(* IEC 61131-3 sources: Lasal-MCP/examples/SampleSource/LASALScreenAdvancedSolution/LASALScreenAdvancedSolution/LASALScreenAdvacnedSolution/Stations/Terminal/HMI/Network/ValueNet, 1 file *)

(* ---- ONE_ValueNet_Table.st ---- *)
#define OBJECTS_CONFIG

FUNCTION GLOBAL TAB ONE_ValueNet
-1$UINT, 0$UINT,
0$UINT, 0$UINT,

1$UDINT,
TO_UDINT(443191026), "MyValues", 0$UINT, 0$UINT, 20$UINT,

_NO_ATTR, TO_UDINT(3497334281), "MYVALUES1",
_NO_ATTR, TO_UDINT(2379682451), "MYVALUES10",
_NO_ATTR, TO_UDINT(4207944197), "MYVALUES11",
_NO_ATTR, TO_UDINT(1675195327), "MYVALUES12",
_NO_ATTR, TO_UDINT(350110505), "MYVALUES13",
_NO_ATTR, TO_UDINT(2327500426), "MYVALUES14",
_NO_ATTR, TO_UDINT(4257080860), "MYVALUES15",
_NO_ATTR, TO_UDINT(1689565094), "MYVALUES16",
_NO_ATTR, TO_UDINT(330532656), "MYVALUES17",
_NO_ATTR, TO_UDINT(2198641313), "MYVALUES18",
_NO_ATTR, TO_UDINT(4094405175), "MYVALUES19",
_NO_ATTR, TO_UDINT(1232881587), "MYVALUES2",
_NO_ATTR, TO_UDINT(2801418576), "MYVALUES20",
_NO_ATTR, TO_UDINT(1048278821), "MYVALUES3",
_NO_ATTR, TO_UDINT(2686444166), "MYVALUES4",
_NO_ATTR, TO_UDINT(3608728080), "MYVALUES5",
_NO_ATTR, TO_UDINT(1309770666), "MYVALUES6",
_NO_ATTR, TO_UDINT(957788988), "MYVALUES7",
_NO_ATTR, TO_UDINT(2846469805), "MYVALUES8",
_NO_ATTR, TO_UDINT(3735985723), "MYVALUES9",

//Internal connections
0$UDINT,
0$UDINT,
0$UDINT,
0$UDINT,

//Initialization values
0$UDINT,
100$UDINT,
TO_UDINT(0), "", TO_UDINT(111),//|ValueNet.MyValues1.Value1;
TO_UDINT(0), "Value2", TO_UDINT(222),//|ValueNet.MyValues1.Value2;
TO_UDINT(0), "Value3", TO_UDINT(333),//|ValueNet.MyValues1.Value3;
TO_UDINT(0), "Active", TO_UDINT(1),//|ValueNet.MyValues1.Active;
TO_UDINT(0), "ID", TO_UDINT(1),//|ValueNet.MyValues1.ID;
TO_UDINT(1), "", TO_UDINT(111),//|ValueNet.MyValues10.Value1;
TO_UDINT(1), "Value2", TO_UDINT(222),//|ValueNet.MyValues10.Value2;
TO_UDINT(1), "Value3", TO_UDINT(333),//|ValueNet.MyValues10.Value3;
TO_UDINT(1), "Active", TO_UDINT(1),//|ValueNet.MyValues10.Active;
TO_UDINT(1), "ID", TO_UDINT(10),//|ValueNet.MyValues10.ID;
TO_UDINT(2), "", TO_UDINT(111),//|ValueNet.MyValues11.Value1;
TO_UDINT(2), "Value2", TO_UDINT(222),//|ValueNet.MyValues11.Value2;
TO_UDINT(2), "Value3", TO_UDINT(333),//|ValueNet.MyValues11.Value3;
TO_UDINT(2), "Active", TO_UDINT(1),//|ValueNet.MyValues11.Active;
TO_UDINT(2), "ID", TO_UDINT(11),//|ValueNet.MyValues11.ID;
TO_UDINT(3), "", TO_UDINT(111),//|ValueNet.MyValues12.Value1;
TO_UDINT(3), "Value2", TO_UDINT(222),//|ValueNet.MyValues12.Value2;
TO_UDINT(3), "Value3", TO_UDINT(333),//|ValueNet.MyValues12.Value3;
TO_UDINT(3), "Active", TO_UDINT(1),//|ValueNet.MyValues12.Active;
TO_UDINT(3), "ID", TO_UDINT(12),//|ValueNet.MyValues12.ID;
TO_UDINT(4), "", TO_UDINT(111),//|ValueNet.MyValues13.Value1;
TO_UDINT(4), "Value2", TO_UDINT(222),//|ValueNet.MyValues13.Value2;
TO_UDINT(4), "Value3", TO_UDINT(333),//|ValueNet.MyValues13.Value3;
TO_UDINT(4), "Active", TO_UDINT(1),//|ValueNet.MyValues13.Active;
TO_UDINT(4), "ID", TO_UDINT(13),//|ValueNet.MyValues13.ID;
TO_UDINT(5), "", TO_UDINT(111),//|ValueNet.MyValues14.Value1;
TO_UDINT(5), "Value2", TO_UDINT(222),//|ValueNet.MyValues14.Value2;
TO_UDINT(5), "Value3", TO_UDINT(333),//|ValueNet.MyValues14.Value3;
TO_UDINT(5), "Active", TO_UDINT(1),//|ValueNet.MyValues14.Active;
TO_UDINT(5), "ID", TO_UDINT(14),//|ValueNet.MyValues14.ID;
TO_UDINT(6), "", TO_UDINT(111),//|ValueNet.MyValues15.Value1;
TO_UDINT(6), "Value2", TO_UDINT(222),//|ValueNet.MyValues15.Value2;
TO_UDINT(6), "Value3", TO_UDINT(333),//|ValueNet.MyValues15.Value3;
TO_UDINT(6), "Active", TO_UDINT(1),//|ValueNet.MyValues15.Active;
TO_UDINT(6), "ID", TO_UDINT(15),//|ValueNet.MyValues15.ID;
TO_UDINT(7), "", TO_UDINT(111),//|ValueNet.MyValues16.Value1;
TO_UDINT(7), "Value2", TO_UDINT(222),//|ValueNet.MyValues16.Value2;
TO_UDINT(7), "Value3", TO_UDINT(333),//|ValueNet.MyValues16.Value3;
TO_UDINT(7), "Active", TO_UDINT(1),//|ValueNet.MyValues16.Active;
TO_UDINT(7), "ID", TO_UDINT(16),//|ValueNet.MyValues16.ID;
TO_UDINT(8), "", TO_UDINT(111),//|ValueNet.MyValues17.Value1;
TO_UDINT(8), "Value2", TO_UDINT(222),//|ValueNet.MyValues17.Value2;
TO_UDINT(8), "Value3", TO_UDINT(333),//|ValueNet.MyValues17.Value3;
TO_UDINT(8), "Active", TO_UDINT(1),//|ValueNet.MyValues17.Active;
TO_UDINT(8), "ID", TO_UDINT(17),//|ValueNet.MyValues17.ID;
TO_UDINT(9), "", TO_UDINT(111),//|ValueNet.MyValues18.Value1;
TO_UDINT(9), "Value2", TO_UDINT(222),//|ValueNet.MyValues18.Value2;
TO_UDINT(9), "Value3", TO_UDINT(333),//|ValueNet.MyValues18.Value3;
TO_UDINT(9), "Active", TO_UDINT(1),//|ValueNet.MyValues18.Active;
TO_UDINT(9), "ID", TO_UDINT(18),//|ValueNet.MyValues18.ID;
TO_UDINT(10), "", TO_UDINT(111),//|ValueNet.MyValues19.Value1;
TO_UDINT(10), "Value2", TO_UDINT(222),//|ValueNet.MyValues19.Value2;
TO_UDINT(10), "Value3", TO_UDINT(333),//|ValueNet.MyValues19.Value3;
TO_UDINT(10), "Active", TO_UDINT(1),//|ValueNet.MyValues19.Active;
TO_UDINT(10), "ID", TO_UDINT(19),//|ValueNet.MyValues19.ID;
TO_UDINT(11), "", TO_UDINT(111),//|ValueNet.MyValues2.Value1;
TO_UDINT(11), "Value2", TO_UDINT(222),//|ValueNet.MyValues2.Value2;
TO_UDINT(11), "Value3", TO_UDINT(333),//|ValueNet.MyValues2.Value3;
TO_UDINT(11), "Active", TO_UDINT(1),//|ValueNet.MyValues2.Active;
TO_UDINT(11), "ID", TO_UDINT(2),//|ValueNet.MyValues2.ID;
TO_UDINT(12), "", TO_UDINT(111),//|ValueNet.MyValues20.Value1;
TO_UDINT(12), "Value2", TO_UDINT(222),//|ValueNet.MyValues20.Value2;
TO_UDINT(12), "Value3", TO_UDINT(333),//|ValueNet.MyValues20.Value3;
TO_UDINT(12), "Active", TO_UDINT(1),//|ValueNet.MyValues20.Active;
TO_UDINT(12), "ID", TO_UDINT(20),//|ValueNet.MyValues20.ID;
TO_UDINT(13), "", TO_UDINT(111),//|ValueNet.MyValues3.Value1;
TO_UDINT(13), "Value2", TO_UDINT(222),//|ValueNet.MyValues3.Value2;
TO_UDINT(13), "Value3", TO_UDINT(333),//|ValueNet.MyValues3.Value3;
TO_UDINT(13), "Active", TO_UDINT(1),//|ValueNet.MyValues3.Active;
TO_UDINT(13), "ID", TO_UDINT(3),//|ValueNet.MyValues3.ID;
TO_UDINT(14), "", TO_UDINT(111),//|ValueNet.MyValues4.Value1;
TO_UDINT(14), "Value2", TO_UDINT(222),//|ValueNet.MyValues4.Value2;
TO_UDINT(14), "Value3", TO_UDINT(333),//|ValueNet.MyValues4.Value3;
TO_UDINT(14), "Active", TO_UDINT(1),//|ValueNet.MyValues4.Active;
TO_UDINT(14), "ID", TO_UDINT(4),//|ValueNet.MyValues4.ID;
TO_UDINT(15), "", TO_UDINT(111),//|ValueNet.MyValues5.Value1;
TO_UDINT(15), "Value2", TO_UDINT(222),//|ValueNet.MyValues5.Value2;
TO_UDINT(15), "Value3", TO_UDINT(333),//|ValueNet.MyValues5.Value3;
TO_UDINT(15), "Active", TO_UDINT(1),//|ValueNet.MyValues5.Active;
TO_UDINT(15), "ID", TO_UDINT(5),//|ValueNet.MyValues5.ID;
TO_UDINT(16), "", TO_UDINT(111),//|ValueNet.MyValues6.Value1;
TO_UDINT(16), "Value2", TO_UDINT(222),//|ValueNet.MyValues6.Value2;
TO_UDINT(16), "Value3", TO_UDINT(333),//|ValueNet.MyValues6.Value3;
TO_UDINT(16), "Active", TO_UDINT(1),//|ValueNet.MyValues6.Active;
TO_UDINT(16), "ID", TO_UDINT(6),//|ValueNet.MyValues6.ID;
TO_UDINT(17), "", TO_UDINT(111),//|ValueNet.MyValues7.Value1;
TO_UDINT(17), "Value2", TO_UDINT(222),//|ValueNet.MyValues7.Value2;
TO_UDINT(17), "Value3", TO_UDINT(333),//|ValueNet.MyValues7.Value3;
TO_UDINT(17), "Active", TO_UDINT(1),//|ValueNet.MyValues7.Active;
TO_UDINT(17), "ID", TO_UDINT(7),//|ValueNet.MyValues7.ID;
TO_UDINT(18), "", TO_UDINT(111),//|ValueNet.MyValues8.Value1;
TO_UDINT(18), "Value2", TO_UDINT(222),//|ValueNet.MyValues8.Value2;
TO_UDINT(18), "Value3", TO_UDINT(333),//|ValueNet.MyValues8.Value3;
TO_UDINT(18), "Active", TO_UDINT(1),//|ValueNet.MyValues8.Active;
TO_UDINT(18), "ID", TO_UDINT(8),//|ValueNet.MyValues8.ID;
TO_UDINT(19), "", TO_UDINT(111),//|ValueNet.MyValues9.Value1;
TO_UDINT(19), "Value2", TO_UDINT(222),//|ValueNet.MyValues9.Value2;
TO_UDINT(19), "Value3", TO_UDINT(333),//|ValueNet.MyValues9.Value3;
TO_UDINT(19), "Active", TO_UDINT(1),//|ValueNet.MyValues9.Active;
TO_UDINT(19), "ID", TO_UDINT(9),//|ValueNet.MyValues9.ID;

//Symbolic initialization values
0$UDINT,
0$UDINT,

//Initialization of string values
0$UDINT,
0$UDINT,

//Configuration of tasks (RealTime, Cyclic, Background)
0$UDINT,
0$UDINT,

0$UDINT,
0$UDINT,

0$UDINT,
0$UDINT,

//External connections
0$UDINT,
0$UDINT,

//Magic internal connections
0$UDINT,
0$UDINT,

//Configuration of timeslots of tasks (RealTime, Cyclic)
#ifdef __LSLLDR_TIMESLOTS__
0$UDINT,
0$UDINT,

0$UDINT,
0$UDINT,

#endif //__LSLLDR_TIMESLOTS__

//MultiMaster connections
#ifdef __LSLLDR_MULTIMASTER__
0$UDINT,
0$UDINT,
#endif //__LSLLDR_MULTIMASTER__

//Configuration for task ID (RealTime, CyclicTime)
#ifdef __LSLLDR_TASKID__
"\\\\TASKS2  "
0$UDINT,
0$UDINT,

0$UDINT,
0$UDINT,

0$UDINT,
0$UDINT,

#endif //__LSLLDR_TASKID__

END_FUNCTION
